TYPE ST_Piston_U_L :
STRUCT
	exist		: 	BOOL	; // true if device exist
	bError		:	BOOL	;
	iFB_Num		: E_Pis_Name;//Parent valve ID number

	//request
	req_Open	:	BOOL	;
	req_Close	:	BOOL	;
	req_Upper	:	BOOL	;
	req_Lower	:	BOOL	;
	req_None		:	BOOL	;
	
	//status
	st_Upper		:	BOOL	;
	st_Lower		:	BOOL	;
	st_Released		:	BOOL	;
	
	
	//Output
	out_Lower	:	BOOL	;
	out_Upper	:	BOOL	;
	
	//sensors
	sen_Upper			:	BOOL	;
	sen_Lower			:	BOOL	;	
	sen_Upper_exist		:	BOOL	;
	sen_Lower_exist		:	BOOL	;	
	//getting the structure of piston
	//str_Piston	:	REFERENCE TO ST_Piston	;
END_STRUCT
END_TYPE

(* stored: Version 1.1.0.1, ProductVersion 3.1.4024.13
   DUT ST_Piston_U_L: Id {b9eedc0d-0f21-48c9-bd0f-9c836f73c0a0} *)
